// TIA Portal V20 export
// export: Created 2026-10-12T15:48:31.7630591Z, ExportSetting WithDefaults, DisplayName Totally Integrated Automation Portal, DisplayVersion V20, DisplayName TIA Portal Openness, DisplayVersion V20, DisplayName TIA Portal Teamcenter Gateway, DisplayVersion V20, DisplayName TIA Portal Version Control Interface, DisplayVersion V20, DisplayName SINAMICS Startdrive Advanced, DisplayVersion V20 SP1 Update 2, DisplayName SINAMICS Startdrive G110M, G120, G120C, G120D, G120P, G115D, DisplayVersion V20 SP1 Update 2, DisplayName SINAMICS Startdrive G130, G150, S120, S150, SINAMICS MV, G220, S200, S210, DisplayVersion V20 SP1 Update 2, DisplayName STEP 7 Professional, DisplayVersion V20, DisplayName STEP 7 Safety, DisplayVersion V20, DisplayName WinCC Basic/Comfort/Advanced, DisplayVersion V20, DisplayName WinCC Professional, DisplayVersion V20, DisplayName WinCC Unified, DisplayVersion V20
FUNCTION "FRK_AlarmHistoryHeaderCrc" : DWord   // FC42, SCL
{ S7_Optimized_Access := 'TRUE' }
VERSION : 0.1
// stored: AutoNumber true, IsIECCheckEnabled false, SetENOAutomatically false, UDAEnableTagReadback false
   VAR_INPUT
      Slot : Int;
   END_VAR
   VAR_TEMP
      Work : DWord;
      Index : Int;
      Size : Int;
   END_VAR
BEGIN

   #FRK_AlarmHistoryHeaderCrc := DWORD#0;
   IF #Slot < 1 OR #Slot > 3 THEN
       RETURN;
   END_IF;
   #Work := "FRK_CrcNumber"(Previous := DWORD#16#FFFFFFFF,
                            Value := UINT_TO_UDINT("FRK_AlarmHistory".Rows[#Slot].SchemaVersion));
   #Size := LEN("FRK_AlarmHistory".Rows[#Slot].Scope);
   #Work := "FRK_CrcNumber"(Previous := #Work,
                            Value := INT_TO_UDINT(#Size));
   FOR #Index := 1 TO #Size DO
       #Work := "FRK_CrcByte"(Previous := #Work,
                              Value := CHAR_TO_BYTE("FRK_AlarmHistory".Rows[#Slot].Scope[#Index]));
   END_FOR;
   #Work := "FRK_CrcNumber"(Previous := #Work,
                            Value := "FRK_AlarmHistory".Rows[#Slot].Generation);
   #Work := "FRK_CrcNumber"(Previous := #Work,
                            Value := INT_TO_UDINT("FRK_AlarmHistory".Rows[#Slot].RingHead));
   #Work := "FRK_CrcNumber"(Previous := #Work,
                            Value := INT_TO_UDINT("FRK_AlarmHistory".Rows[#Slot].RingUsed));
   #Work := "FRK_CrcNumber"(Previous := #Work,
                            Value := BOOL_TO_UDINT("FRK_AlarmHistory".Rows[#Slot].Truncated));
   FOR #Index := 1 TO 64 DO
       #Work := "FRK_CrcNumber"(Previous := #Work,
                                Value := DWORD_TO_UDINT("FRK_AlarmHistory".Rows[#Slot].EventCrc[#Index]));
   END_FOR;
   #FRK_AlarmHistoryHeaderCrc := NOT #Work;
END_FUNCTION
